// TIA Portal V19 export
DATA_BLOCK "ALL_VALVES_DB"   // DB14
// stored: InstanceOfName ALL_VALVES, InstanceOfType FB
"ALL_VALVES"
   // VAR
   //    valve_R1_XV01 { S7_SetPoint := 'True'} : "valve";
   //    valve_R1_XV02 { S7_SetPoint := 'True'} : "valve";
   //    valve_R1_XV03 { S7_SetPoint := 'True'} : "valve";
   //    valve_R1_XV04 { S7_SetPoint := 'True'} : "valve";
   //    valve_R1_XV05 { S7_SetPoint := 'True'} : "valve";
   //    valve_R1_XV06 { S7_SetPoint := 'True'} : "valve";
   //    valve_R1_XV07 { S7_SetPoint := 'True'} : "valve";
   //    valve_R1_XV08 { S7_SetPoint := 'True'} : "valve";
   //    valve_R1_XV09 { S7_SetPoint := 'True'} : "valve";
   //    valve_R1_XV10 { S7_SetPoint := 'True'} : "valve";
   //    clod_skid { S7_SetPoint := 'True'} : "valve";
   //    valve_R2_XV01 { S7_SetPoint := 'True'} : "valve";
   //    valve_R2_XV02 { S7_SetPoint := 'True'} : "valve";
   //    valve_R2_XV03 { S7_SetPoint := 'True'} : "valve";
   //    valve_R2_XV04 { S7_SetPoint := 'True'} : "valve";
   //    valve_R2_XV05 { S7_SetPoint := 'True'} : "valve";
   //    valve_R2_XV06 { S7_SetPoint := 'True'} : "valve";
   //    valve_R2_XV07 { S7_SetPoint := 'True'} : "valve";
   //    valve_R2_XV08 { S7_SetPoint := 'True'} : "valve";
   //    valve_R2_XV09 { S7_SetPoint := 'True'} : "valve";
   //    valve_R2_XV10 { S7_SetPoint := 'True'} : "valve";
   //    valve_R3_XV01 { S7_SetPoint := 'True'} : "valve";
   //    valve_R3_XV02 { S7_SetPoint := 'True'} : "valve";
   //    valve_R3_XV03 { S7_SetPoint := 'True'} : "valve";
   //    valve_R3_XV04 { S7_SetPoint := 'True'} : "valve";
   //    valve_R3_XV05 { S7_SetPoint := 'True'} : "valve";
   //    valve_R3_XV06 { S7_SetPoint := 'True'} : "valve";
   //    valve_R3_XV07 { S7_SetPoint := 'True'} : "valve";
   //    valve_R3_XV08 { S7_SetPoint := 'True'} : "valve";
   //    valve_R3_XV09 { S7_SetPoint := 'True'} : "valve";
   //    valve_R3_XV10 { S7_SetPoint := 'True'} : "valve";
   //    valve_R4_XV02 { S7_SetPoint := 'True'} : "valve";
   //    valve_R4_XV01 { S7_SetPoint := 'True'} : "valve";
   //    valve_R4_XV03 { S7_SetPoint := 'True'} : "valve";
   //    valve_R4_XV04 { S7_SetPoint := 'True'} : "valve";
   //    valve_R4_XV05 { S7_SetPoint := 'True'} : "valve";
   //    valve_R4_XV06 { S7_SetPoint := 'True'} : "valve";
   //    valve_R4_XV07 { S7_SetPoint := 'True'} : "valve";
   //    valve_R4_XV08 { S7_SetPoint := 'True'} : "valve";
   //    valve_R4_XV09 { S7_SetPoint := 'True'} : "valve";
   //    valve_R4_XV10 { S7_SetPoint := 'True'} : "valve";
   //    valve_R8_XV2 { S7_SetPoint := 'True'} : "valve";
   //    valve_R8_XV3 { S7_SetPoint := 'True'} : "valve";
   //    valve_R8_XV4 { S7_SetPoint := 'True'} : "valve";
   //    valve_R8_XV5 { S7_SetPoint := 'True'} : "valve";
   //    valve_R8_XV05 { S7_SetPoint := 'True'} : "valve";
   //    valve_R8_XV06 { S7_SetPoint := 'True'} : "valve";
   //    valve_R8_XV07 { S7_SetPoint := 'True'} : "valve";
   //    valve_R8_XV08 { S7_SetPoint := 'True'} : "valve";
   //    valve_R8_XV09 { S7_SetPoint := 'True'} : "valve";
   //    valve_R8_XV10 { S7_SetPoint := 'True'} : "valve";
   //    valve_R6_XV01 { S7_SetPoint := 'True'} : "valve";
   //    valve_R6_XV02 { S7_SetPoint := 'True'} : "valve";
   //    valve_R6_XV03 { S7_SetPoint := 'True'} : "valve";
   //    valve_R6_XV04 { S7_SetPoint := 'True'} : "valve";
   //    valve_R6_XV05 { S7_SetPoint := 'True'} : "valve";
   //    valve_R6_XV06 { S7_SetPoint := 'True'} : "valve";
   //    valve_R6_XV07 { S7_SetPoint := 'True'} : "valve";
   //    valve_R6_XV08 { S7_SetPoint := 'True'} : "valve";
   //    valve_R6_XV09 { S7_SetPoint := 'True'} : "valve";
   //    valve_R6_XV10 { S7_SetPoint := 'True'} : "valve";
   //    valve_R7_XV01 { S7_SetPoint := 'True'} : "valve";
   //    valve_R7_XV02 { S7_SetPoint := 'True'} : "valve";
   //    valve_R7_XV03 { S7_SetPoint := 'True'} : "valve";
   //    valve_R7_XV04 { S7_SetPoint := 'True'} : "valve";
   //    valve_R7_XV05 { S7_SetPoint := 'True'} : "valve";
   //    valve_R7_XV06 { S7_SetPoint := 'True'} : "valve";
   //    valve_R7_XV07 { S7_SetPoint := 'True'} : "valve";
   //    valve_R7_XV08 { S7_SetPoint := 'True'} : "valve";
   //    valve_R7_XV09 { S7_SetPoint := 'True'} : "valve";
   //    valve_R7_XV10 { S7_SetPoint := 'True'} : "valve";
   //    valve_R8_XV01 { S7_SetPoint := 'True'} : "valve";
   //    valve_R8_XV02 { S7_SetPoint := 'True'} : "valve";
   //    valve_R8_XV03 { S7_SetPoint := 'True'} : "valve";
   //    valve_R8_XV04 { S7_SetPoint := 'True'} : "valve";
   //    valve_R5_XV2 { S7_SetPoint := 'True'} : "valve";
   //    valve_R5_XV3 { S7_SetPoint := 'True'} : "valve";
   //    valve_R5_XV4 { S7_SetPoint := 'True'} : "valve";
   //    valve_R5_XV5 { S7_SetPoint := 'True'} : "valve";
   //    valve_R5_XV05 { S7_SetPoint := 'True'} : "valve";
   //    valve_R5_XV06 { S7_SetPoint := 'True'} : "valve";
   //    valve_R5_XV07 { S7_SetPoint := 'True'} : "valve";
   //    valve_R5_XV08 { S7_SetPoint := 'True'} : "valve";
   //    valve_R5_XV09 { S7_SetPoint := 'True'} : "valve";
   //    valve_R5_XV10 { S7_SetPoint := 'True'} : "valve";
   //    valve_R9_XV01 { S7_SetPoint := 'True'} : "valve";
   //    valve_R9_XV02 { S7_SetPoint := 'True'} : "valve";
   //    valve_R9_XV03 { S7_SetPoint := 'True'} : "valve";
   //    valve_R9_XV04 { S7_SetPoint := 'True'} : "valve";
   //    valve_R9_XV05 { S7_SetPoint := 'True'} : "valve";
   //    valve_R9_XV06 { S7_SetPoint := 'True'} : "valve";
   //    valve_R9_XV07 { S7_SetPoint := 'True'} : "valve";
   //    valve_R9_XV08 { S7_SetPoint := 'True'} : "valve";
   //    valve_R9_XV09 { S7_SetPoint := 'True'} : "valve";
   //    valve_R9_XV10 { S7_SetPoint := 'True'} : "valve";
   //    valve_R10_XV01 { S7_SetPoint := 'True'} : "valve";
   //    valve_R10_XV02 { S7_SetPoint := 'True'} : "valve";
   //    valve_R10_XV03 { S7_SetPoint := 'True'} : "valve";
   //    valve_R10_XV04 { S7_SetPoint := 'True'} : "valve";
   //    valve_R10_XV05 { S7_SetPoint := 'True'} : "valve";
   //    valve_R10_XV06 { S7_SetPoint := 'True'} : "valve";
   //    valve_R10_XV07 { S7_SetPoint := 'True'} : "valve";
   //    valve_R10_XV08 { S7_SetPoint := 'True'} : "valve";
   //    valve_R10_XV09 { S7_SetPoint := 'True'} : "valve";
   //    valve_R10_XV10 { S7_SetPoint := 'True'} : "valve";
   //    valve_R11_XV01 { S7_SetPoint := 'True'} : "valve";
   //    valve_R11_XV02 { S7_SetPoint := 'True'} : "valve";
   //    valve_R11_XV03 { S7_SetPoint := 'True'} : "valve";
   //    valve_R11_XV04 { S7_SetPoint := 'True'} : "valve";
   //    valve_R11_XV05 { S7_SetPoint := 'True'} : "valve";
   //    valve_R11_XV06 { S7_SetPoint := 'True'} : "valve";
   //    valve_R11_XV07 { S7_SetPoint := 'True'} : "valve";
   //    valve_R11_XV08 { S7_SetPoint := 'True'} : "valve";
   //    valve_R11_XV09 { S7_SetPoint := 'True'} : "valve";
   //    valve_R11_XV10 { S7_SetPoint := 'True'} : "valve";
   //    valve_R12_XV01 { S7_SetPoint := 'True'} : "valve";
   //    valve_R12_XV02 { S7_SetPoint := 'True'} : "valve";
   //    valve_R12_XV03 { S7_SetPoint := 'True'} : "valve";
   //    valve_R12_XV04 { S7_SetPoint := 'True'} : "valve";
   //    valve_R12_XV05 { S7_SetPoint := 'True'} : "valve";
   //    valve_R12_XV06 { S7_SetPoint := 'True'} : "valve";
   //    valve_R12_XV07 { S7_SetPoint := 'True'} : "valve";
   //    valve_R12_XV08 { S7_SetPoint := 'True'} : "valve";
   //    valve_R12_XV09 { S7_SetPoint := 'True'} : "valve";
   //    valve_R12_XV10 { S7_SetPoint := 'True'} : "valve";
   //    valve_R13_XV01 { S7_SetPoint := 'True'} : "valve";
   //    valve_R13_XV02 { S7_SetPoint := 'True'} : "valve";
   //    valve_R13_XV03 { S7_SetPoint := 'True'} : "valve";
   //    valve_R13_XV04 { S7_SetPoint := 'True'} : "valve";
   //    valve_R13_XV05 { S7_SetPoint := 'True'} : "valve";
   //    valve_R13_XV06 { S7_SetPoint := 'True'} : "valve";
   //    valve_R13_XV07 { S7_SetPoint := 'True'} : "valve";
   //    valve_R13_XV08 { S7_SetPoint := 'True'} : "valve";
   //    valve_R13_XV09 { S7_SetPoint := 'True'} : "valve";
   //    valve_R13_XV10 { S7_SetPoint := 'True'} : "valve";
   //    valve_R14_XV02 { S7_SetPoint := 'True'} : "valve";
   //    valve_R14_XV01 { S7_SetPoint := 'True'} : "valve";
   //    valve_R14_XV03 { S7_SetPoint := 'True'} : "valve";
   //    valve_R14_XV04 { S7_SetPoint := 'True'} : "valve";
   //    valve_R14_XV05 { S7_SetPoint := 'True'} : "valve";
   //    valve_R14_XV06 { S7_SetPoint := 'True'} : "valve";
   //    valve_R14_XV07 { S7_SetPoint := 'True'} : "valve";
   //    valve_R14_XV08 { S7_SetPoint := 'True'} : "valve";
   //    valve_R14_XV09 { S7_SetPoint := 'True'} : "valve";
   //    valve_R14_XV10 { S7_SetPoint := 'True'} : "valve";
   //    valve_R15_XV02 { S7_SetPoint := 'True'} : "valve";
   //    valve_R15_XV01 { S7_SetPoint := 'True'} : "valve";
   //    valve_R15_XV03 { S7_SetPoint := 'True'} : "valve";
   //    valve_R15_XV04 { S7_SetPoint := 'True'} : "valve";
   //    valve_R15_XV05 { S7_SetPoint := 'True'} : "valve";
   //    valve_R15_XV06 { S7_SetPoint := 'True'} : "valve";
   //    valve_R15_XV07 { S7_SetPoint := 'True'} : "valve";
   //    valve_R15_XV08 { S7_SetPoint := 'True'} : "valve";
   //    valve_R15_XV09 { S7_SetPoint := 'True'} : "valve";
   //    valve_R15_XV10 { S7_SetPoint := 'True'} : "valve";
   //    valve_R16_XV02 { S7_SetPoint := 'True'} : "valve";
   //    valve_R16_XV03 { S7_SetPoint := 'True'} : "valve";
   //    valve_R16_XV04 { S7_SetPoint := 'True'} : "valve";
   //    valve_R16_XV05 { S7_SetPoint := 'True'} : "valve";
   //    valve_R16_XV06 { S7_SetPoint := 'True'} : "valve";
   //    valve_R16_XV07 { S7_SetPoint := 'True'} : "valve";
   //    valve_R16_XV08 { S7_SetPoint := 'True'} : "valve";
   //    valve_R16_XV09 { S7_SetPoint := 'True'} : "valve";
   //    valve_R16_XV10 { S7_SetPoint := 'True'} : "valve";
   //    valve_R17_XV01 { S7_SetPoint := 'True'} : "valve";
   //    valve_R17_XV02 { S7_SetPoint := 'True'} : "valve";
   //    valve_R17_XV03 { S7_SetPoint := 'True'} : "valve";
   //    valve_R17_XV04 { S7_SetPoint := 'True'} : "valve";
   //    valve_R17_XV05 { S7_SetPoint := 'True'} : "valve";
   //    valve_R17_XV06 { S7_SetPoint := 'True'} : "valve";
   //    valve_R17_XV07 { S7_SetPoint := 'True'} : "valve";
   //    valve_R17_XV08 { S7_SetPoint := 'True'} : "valve";
   //    valve_R17_XV09 { S7_SetPoint := 'True'} : "valve";
   //    valve_R17_XV10 { S7_SetPoint := 'True'} : "valve";
   //    valve_R18_XV02 { S7_SetPoint := 'True'} : "valve";
   //    valve_R18_XV03 { S7_SetPoint := 'True'} : "valve";
   //    valve_R18_XV04 { S7_SetPoint := 'True'} : "valve";
   //    valve_R18_XV05 { S7_SetPoint := 'True'} : "valve";
   //    valve_R18_XV06 { S7_SetPoint := 'True'} : "valve";
   //    valve_R18_XV07 { S7_SetPoint := 'True'} : "valve";
   //    valve_R18_XV08 { S7_SetPoint := 'True'} : "valve";
   //    valve_R18_XV09 { S7_SetPoint := 'True'} : "valve";
   //    valve_R18_XV10 { S7_SetPoint := 'True'} : "valve";
   //    child_skid { S7_SetPoint := 'True'} : "valve";
   //    ultra_child { S7_SetPoint := 'True'} : "valve";
   // END_VAR
BEGIN
END_DATA_BLOCK
